// TIA Portal V19 export
TYPE "Pan_To_SM"
   STRUCT
      Massecuite_Solids : Real;
      Level : Real;
      Absolute_Pressure : Real;
      Purity_P1 : Real;
      Purity_P2 : Real;
      Purity_P3 : Real;
      Purity_Selector : UInt;
      Final_Mass_Solid_Prog1 : Real;
      Final_Mass_Solid_Prog2 : Real;
      Final_Mass_Solid_Prog3 : Real;
      Final_Mass_Solid_Selector : UInt;
      Strike_Active : Bool;
      Seeded : Bool;
      reserve_bit_2 : Bool;
      SM_Auto_Seeding_Required : Bool;
      reserve_bit_4 : Bool;
      reserve_bit_5 : Bool;
      reserve_bit_6 : Bool;
      reserve_bit_7 : Bool;
   END_STRUCT;
END_TYPE
